Staubli VAL3: utCommon.dtx

public bool bDisabled
public string sValue
public string sID
public num nValue
public string sPage
